(* IEC 61131-3 sources: test/Class/SdiasSDCIMaster (part 4) *)

          GetSdoReadData(pLength:=#TempDataLen, pData:=#TempData[0]);
          if TempDataLen = 9 then
            // check response data
            if (TempData[0] = (E_FNCID_CNTSTA)$USINT) then // check function ID
              // reset response state machine
              sSdoData.eResponseState := t_ReponseState::_PrepareSendData;

              // if the operating flags are cleared we can continue
              for i:= 0 to SIOL_MAX_PORTS_SUPPORTED-1 do
                TempStateFlags := TempData[1 + i*sizeof(t_StatusFlags)]$t_StatusFlags;

                // if any operating bit of the SDCI ports is still set and we did not exceed the timeout => go to wait for disabled
                if (aPortInfo[i].CfgPortMode = _SDCI) & (TempStateFlags.Operating = TRUE) &
                   ((ops.tAbsolute - Wait4DeviceDisableStartTime) < aPortInfo[sSdoData.ActPortSelection].udModeChangeTime) then

                  sSdoData.eInitSSW   := t_InitSSW::_Wait4DisableMode2;
                  return;
                end_if;
              end_for;

              // finished, continue with next step
              sSdoData.eInitSSW   := t_InitSSW::_Configure2StartUpMode;

            else
              // unexpected answer data
              LogError("@0525 (SdiasSDCIMaster::InitTheModule) Unexpected data in answer from µC: wrong function ID or port number (_SwitchToDisableMode2)");
              sSdoData.eInitSSW := _Error;
              return;
            end_if;
          else
            // invalid length of answer data
            LogError("@0526 (SdiasSDCIMaster::InitTheModule) Invalid data length in answer from µC (_SwitchToDisableMode2)");
            sSdoData.eInitSSW := _Error;
            return;
          end_if;

      //***************************************************************************************************
      end_case;

//**********************************************************************************************************************************************************
  	t_InitSSW::_Configure2StartUpMode:
      // if it's an SDCI port and physically available, we must wait the time (according to the specification), because some sensors might need it
      if (aPortInfo[sSdoData.ActPortSelection].CfgPortMode = _SDCI) &
          aPortInfo[sSdoData.ActPortSelection].PhysicallyAvailable  &
         ((ops.tAbsolute - Wait4DeviceDisableStartTime) < aPortInfo[sSdoData.ActPortSelection].udModeChangeTime) then
        return;
      end_if;

      case sSdoData.eResponseState of
      //***************************************************************************************************
        t_ReponseState::_PrepareSendData: // start the sending action

          // only if the port is of type SDCI and the device is physically available
          if (aPortInfo[sSdoData.ActPortSelection].CfgPortMode = _SDCI) & aPortInfo[sSdoData.ActPortSelection].PhysicallyAvailable &
             (aPortInfo[sSdoData.ActPortSelection].StartUpMode <> _Inactive) then

            // prepare the sdo buffer
            TempData[0]       := E_FNCID_SETPORTCNFPAR; // function ID
            TempData[1]       := sSdoData.ActPortSelection; // port number

            case aPortInfo[sSdoData.ActPortSelection].StartUpMode of
            //***************************************************************************************************
              _DigitalInput:
                TempData[2]       := t_OpModeStates::E_OPMODE_DI; // operating mode

            //***************************************************************************************************
              _DigitalOutput:
                TempData[2]       := t_OpModeStates::E_OPMODE_DO; // operating mode

            //***************************************************************************************************
              _SDCI:
                TempData[2]       := t_OpModeStates::E_OPMODE_FIXEDMODE; // operating mode

            //***************************************************************************************************
            end_case;

            TempData[3]       := t_PortCycle::E_PORTCYCLE_FIXVAL; // port cycle

            // check if a user override is active
            if aPortInfo[sSdoData.ActPortSelection].OverrideMinCycleTime_us then
              // recalculate cycle time from [µs] to [100µs]
              TempCycleTime     := to_uint(aPortInfo[sSdoData.ActPortSelection].OverrideMinCycleTime_us / 100);
            else
              // recalculate cycle time from [µs] to [100µs]
              TempCycleTime     := to_uint(aPortInfo[sSdoData.ActPortSelection].MinCycleTime_us / 100);
            end_if;

            // make endian swap
            TempCycleTime     := ((TempCycleTime SHR 8) AND 16#FF) OR ((TempCycleTime SHL 8) AND 16#FF00);

            TempData[4]$UINT  := TempCycleTime; // cycle time
            TempData[6]       :=  aPortInfo[sSdoData.ActPortSelection].PdoMapping.ReadDataLength$USINT; // PDConfig LenIn
            TempData[7]       := (aPortInfo[sSdoData.ActPortSelection].PdoMapping.ReadDataStartAddress - SIOL_OFFSET_RT_READ_DATA)$USINT; // PdConfig PosIn
            TempData[8]       := 0; // PdConfig SrcOffsetIn
            TempData[9]       :=  aPortInfo[sSdoData.ActPortSelection].PdoMapping.WriteDataLength$USINT; // PDConfig LenOut
            TempData[10]      := (aPortInfo[sSdoData.ActPortSelection].PdoMapping.WriteDataStartAddress - SIOL_OFFSET_RT_WRITE_DATA)$USINT; // PdConfig PosOut
            TempData[11]      := 0; // PdConfig SrcOffsetOut
            TempData[12]      := (aPortInfo[sSdoData.ActPortSelection].VendorID SHR 8)$USINT; // VendorID
            TempData[13]      :=  aPortInfo[sSdoData.ActPortSelection].VendorID$USINT; // VendorID
            TempData[14]      := (aPortInfo[sSdoData.ActPortSelection].DeviceID SHR 24)$USINT; // DeviceID
            TempData[15]      := (aPortInfo[sSdoData.ActPortSelection].DeviceID SHR 16)$USINT; // DeviceID
            TempData[16]      := (aPortInfo[sSdoData.ActPortSelection].DeviceID SHR  8)$USINT; // DeviceID
            TempData[17]      := (aPortInfo[sSdoData.ActPortSelection].DeviceID       )$USINT; // DeviceID
  //          _strcpy(dest:=#TempData[18], src:="0000000000000000"); // serial number as string
            _memset(dest:=#TempData[18], usByte:=0, cntr:=16); // serial number as string
            TempData[34]      := 1; // Inspection level (1 = device and vendor id have to match)
            TempData[35]      := 0; // DS activation state
            TempData[36]      := 0; // DS download enable
            TempData[37]      := 0; // DS upload enable
            TempData[38]      := aPortInfo[sSdoData.ActPortSelection].RevisionID; // revision ID

            TempDataLen := 39;

            InitializeSdoWriteData(Usage:=_SendFunctionCode, ParaIndex:=0, ParaSubIndex:=0, PortSelection:=SIOL_MASTER_PORT_NO, LengthOfData:=TempDataLen, pData:=#TempData[0]);

            sSdoData.eResponseState := t_ReponseState::_SendData;
          else
            if (aPortInfo[sSdoData.ActPortSelection].CfgPortMode = _SDCI) & (aPortInfo[sSdoData.ActPortSelection].StartUpMode = _Inactive) &
                aPortInfo[sSdoData.ActPortSelection].PhysicallyAvailable then
              // the current mode is now the startupmode
              aPortInfo[sSdoData.ActPortSelection].ActPortMode := aPortInfo[sSdoData.ActPortSelection].StartUpMode;

              // it's always ok here
              MyPara.aPara[0] := _ClassOk$DINT;

              // vendor ID
              MyPara.aPara[1] := aPortInfo[sSdoData.ActPortSelection].VendorID;

              // device ID
              MyPara.aPara[2] := aPortInfo[sSdoData.ActPortSelection].DeviceID$DINT;

              // minimum cycle time
              // check if a user override is active
              if aPortInfo[sSdoData.ActPortSelection].OverrideMinCycleTime_us then
                MyPara.aPara[3] := aPortInfo[sSdoData.ActPortSelection].OverrideMinCycleTime_us$DINT;
              else
                MyPara.aPara[3] := aPortInfo[sSdoData.ActPortSelection].MinCycleTime_us$DINT;
              end_if;

              // actual port mode is already valid here (no further changes on the setting of this port)
              MyPara.aPara[4] := aPortInfo[sSdoData.ActPortSelection].ActPortMode$DINT;

              aPortInfo[sSdoData.ActPortSelection].pThis^.NewInst(#MyPara, #MyResult);
            end_if;

            // already the last port?
            if sSdoData.ActPortSelection = (SIOL_MAX_PORTS_SUPPORTED-1) then
              // finished, continue with next step
              sSdoData.ActPortSelection := 0;
              DelayedEnablePorts        := 0;
              DigStartUpAvailable       := FALSE;

              for i:= 0 to SIOL_MAX_PORTS_SUPPORTED-1 do
                if (aPortInfo[i].CfgPortMode = _SDCI) & aPortInfo[i].PhysicallyAvailable then
                  if (aPortInfo[i].StartUpMode = _SDCI) then
                    DelayedEnablePorts := DelayedEnablePorts OR (1 SHL i$USINT);
                  elsif (aPortInfo[i].StartUpMode = _DigitalInput) | (aPortInfo[i].StartUpMode = _DigitalOutput) then
                    DigStartUpAvailable := TRUE;
                  end_if;
                end_if;
              end_for;

              if DelayedEnablePorts then
                // block the asynchron communication channel already
                sSdoData.AsyState             := t_SDCIRetCode::SDCI_Busy;
                sSdoData.TargetMode           := _SDCI;
                sSdoData.AsyCmdType           := t_AsyCmdType::DelayedEnable;
                sSdoData.eAsySSW              := t_AsySSW::_StartDelayedEnable;
                DelayedEnablePorts.FirstTime  := TRUE; // this is set to reset the port number on the first entrace in cyclic
              end_if;

              if DigStartUpAvailable then
                sSdoData.eInitSSW   := t_InitSSW::_EnableDigIOStartUpModes;
              else
                sSdoData.eInitSSW   := t_InitSSW::_SetCycleTimes;
              end_if;
            else
              // repeat the steps with the next port
              sSdoData.ActPortSelection += 1;
            end_if;
          end_if;

      //***************************************************************************************************
        t_ReponseState::_SendData,
        t_ReponseState::_Wait4SendResponse,
        t_ReponseState::_GotSendResponse,
        t_ReponseState::_ReadData,
        t_ReponseState::_Wait4ReceiveData,
        t_ReponseState::_GotReceiveData:
          if HandleSdoDataTransfer() = ERROR then
            sSdoData.eInitSSW := _Error;
            return;
          end_if;

      //***************************************************************************************************
        t_ReponseState::_GotAllReceiveData:// we enter this step, when we received the answer with the data

          GetSdoReadData(pLength:=#TempDataLen, pData:=#TempData[0]);
          if TempDataLen = 3 then
            // check response data
            if (TempData[0] = (E_FNCID_SETPORTCNFPAR)$USINT) & // check function ID
               (TempData[1] = sSdoData.ActPortSelection)              // check port number
               then

              if (TempData[2] = 0) then // check status code seperately
                // reset response state machine
                sSdoData.eResponseState := t_ReponseState::_PrepareSendData;

                // already the last port?
                if sSdoData.ActPortSelection = (SIOL_MAX_PORTS_SUPPORTED-1) then
                  // finished, continue with next step
                  sSdoData.ActPortSelection := 0;
                  DelayedEnablePorts        := 0;
                  DigStartUpAvailable       := FALSE;

                  for i:= 0 to SIOL_MAX_PORTS_SUPPORTED-1 do
                    if (aPortInfo[i].StartUpMode = _SDCI) & aPortInfo[i].PhysicallyAvailable then
                      DelayedEnablePorts := DelayedEnablePorts OR (1 SHL i$USINT);
                    elsif (aPortInfo[i].CfgPortMode = _SDCI)         &  aPortInfo[i].PhysicallyAvailable &
                         ((aPortInfo[i].StartUpMode = _DigitalInput) | (aPortInfo[i].StartUpMode = _DigitalOutput)) then
                      DigStartUpAvailable := TRUE;
                    end_if;
                  end_for;

                  if DelayedEnablePorts then
                    // block the asynchron communication channel already
                    sSdoData.AsyState             := t_SDCIRetCode::SDCI_Busy;
                    sSdoData.TargetMode           := _SDCI;
                    sSdoData.AsyCmdType           := t_AsyCmdType::DelayedEnable;
                    sSdoData.eAsySSW              := t_AsySSW::_StartDelayedEnable;
                    DelayedEnablePorts.FirstTime  := TRUE; // this is set to reset the port number on the first entrace in cyclic
                  end_if;

                  if DigStartUpAvailable then
                    sSdoData.eInitSSW   := t_InitSSW::_EnableDigIOStartUpModes;
                  else
                    sSdoData.eInitSSW   := t_InitSSW::_SetCycleTimes;
                  end_if;
                else
                  // repeat the steps with the next port
                  sSdoData.ActPortSelection += 1;
                end_if;
              else
                // error at return code
                LogError("@0527 (SdiasSDCIMaster::InitTheModule) Error at status code in answer from µC (_Configure2StartUpMode)");
                sSdoData.eInitSSW := _Error;
                return;
              end_if;
            else
              // unexpected answer data
              LogError("@0529 (SdiasSDCIMaster::InitTheModule) Unexpected data in answer from µC: wrong function ID or port number (_ReEnableWithFixedMode)");
              sSdoData.eInitSSW := _Error;
              return;
            end_if;
          else
            // invalid length of answer data
            LogError("@052A (SdiasSDCIMaster::InitTheModule) Invalid data length in answer from µC (_Configure2StartUpMode)");
            sSdoData.eInitSSW := _Error;
            return;
          end_if;

      //***************************************************************************************************
      end_case;

//**********************************************************************************************************************************************************
  	t_InitSSW::_EnableDigIOStartUpModes:
      case sSdoData.eResponseState of
      //***************************************************************************************************
        t_ReponseState::_PrepareSendData: // start the sending action
          TempFlags := 0;
          TempFlags.Start2Operate := TRUE;
          TempFlags.OperatingMode := TRUE;

          // prepare the sdo buffer
          TempData[0]       := E_FNCID_CNTSTA; // function ID
          for i:= 0 to SIOL_MAX_PORTS_SUPPORTED-1 do

            // if the startup mode is digin or digout => enable this mode now
            if (aPortInfo[i].CfgPortMode = _SDCI)         &  aPortInfo[i].PhysicallyAvailable &
              ((aPortInfo[i].StartUpMode = _DigitalInput) | (aPortInfo[i].StartUpMode = _DigitalOutput)) then
              TempData[1 + i*sizeof(UINT)]$UINT := TempFlags;
            else
              // otherwise don't do anything at this port
              TempData[1 + i*sizeof(UINT)]$UINT := 0;
            end_if;
          end_for;

          if TotalMappingWriteSize then
            _memset(dest:=#TempData[9], usByte:=0, cntr:=TotalMappingWriteSize);
          end_if;

          TempDataLen := 9 + TotalMappingWriteSize;

          InitializeSdoWriteData(Usage:=_SendFunctionCode, ParaIndex:=0, ParaSubIndex:=0, PortSelection:=SIOL_MASTER_PORT_NO, LengthOfData:=TempDataLen, pData:=#TempData[0]);

          sSdoData.eResponseState := t_ReponseState::_SendData;

      //***************************************************************************************************
        t_ReponseState::_SendData,
        t_ReponseState::_Wait4SendResponse,
        t_ReponseState::_GotSendResponse,
        t_ReponseState::_ReadData,
        t_ReponseState::_Wait4ReceiveData,
        t_ReponseState::_GotReceiveData:
          if HandleSdoDataTransfer() = ERROR then
            sSdoData.eInitSSW := _Error;
            return;
          end_if;

      //***************************************************************************************************
        t_ReponseState::_GotAllReceiveData:// we enter this step, when we received the answer with the data

          GetSdoReadData(pLength:=#TempDataLen, pData:=#TempData[0]);
          if TempDataLen = 9 then

            // reset response state machine
            sSdoData.eResponseState := t_ReponseState::_PrepareSendData;

            // check response data
            if (TempData[0] = (E_FNCID_CNTSTA)$USINT) then // check function ID

              // update the state of the object
              for i:= 0 to SIOL_MAX_PORTS_SUPPORTED-1 do

                // if the startup mode is digin or digout => show classok and current mode
                if (aPortInfo[i].CfgPortMode = _SDCI)         &  aPortInfo[i].PhysicallyAvailable
                & ((aPortInfo[i].StartUpMode = _DigitalInput) | (aPortInfo[i].StartUpMode = _DigitalOutput))
                  then
                  // the current mode is now the startupmode
                  aPortInfo[i].ActPortMode := aPortInfo[i].StartUpMode;

                  // it's always ok here
                  MyPara.aPara[0] := _ClassOk$DINT;

                  // vendor ID
                  MyPara.aPara[1] := aPortInfo[i].VendorID;

                  // device ID
                  MyPara.aPara[2] := aPortInfo[i].DeviceID$DINT;

                  // minimum cycle time
                  // check if a user override is active
                  if aPortInfo[i].OverrideMinCycleTime_us then
                    MyPara.aPara[3] := aPortInfo[i].OverrideMinCycleTime_us$DINT;
                  else
                    MyPara.aPara[3] := aPortInfo[i].MinCycleTime_us$DINT;
                  end_if;

                  // actual port mode is already valid here (no further changes on the setting of this port)
                  MyPara.aPara[4] := aPortInfo[i].ActPortMode$DINT;

                  aPortInfo[i].pThis^.NewInst(#MyPara, #MyResult);
                end_if;
              end_for;

              // finished, continue with next step
              sSdoData.eInitSSW   := t_InitSSW::_SetCycleTimes;

            else
              // unexpected answer data
              LogError("@050C (SdiasSDCIMaster::InitTheModule) Unexpected data in answer from µC: wrong function ID or port number (_SwitchToNewMode)");
              sSdoData.eInitSSW := _Error;
              return;
            end_if;
          else
            // invalid length of answer data
            LogError("@050D (SdiasSDCIMaster::InitTheModule) Invalid data length in answer from µC (_SwitchToNewMode)");
            sSdoData.eInitSSW := _Error;
            return;
          end_if;

      //***************************************************************************************************
      end_case;

//**********************************************************************************************************************************************************
  	t_InitSSW::_SetCycleTimes:

      case sSdoData.eResponseState of
      //***************************************************************************************************
        t_ReponseState::_PrepareSendData: // start the sending action

          // take the time from the parameter download process
          ParaDownloadTime := ops.tAbsolute - DownloadTimeStart;

          TempData[0]$UINT  := (udBusTime / 1000)$UINT; // SDIAS Bus cycle time
          TempData[2]$UINT  := CycleTime$UINT;

          TempDataLen    := 2 * sizeof(UINT);

          InitializeSdoWriteData(Usage:=_SendCycleTimeInfo, ParaIndex:=0, ParaSubIndex:=0, PortSelection:=SIOL_MASTER_PORT_NO, LengthOfData:=TempDataLen, pData:=#TempData[0]);

          sSdoData.eResponseState := t_ReponseState::_SendData;

      //***************************************************************************************************
        t_ReponseState::_SendData,
        t_ReponseState::_Wait4SendResponse,
        t_ReponseState::_GotSendResponse,
        t_ReponseState::_ReadData,
        t_ReponseState::_Wait4ReceiveData,
        t_ReponseState::_GotReceiveData:
          if HandleSdoDataTransfer() = ERROR then
            sSdoData.eInitSSW := _Error;
            return;
          end_if;

      //***************************************************************************************************
        t_ReponseState::_GotAllReceiveData:// we enter this step, when we received the answer with the data

          GetSdoReadData(pLength:=#TempDataLen, pData:=#TempData[0]);
          if TempDataLen = 0 then
            // check response data
            if (sSdoData.SdoReadData.ro_RetCode = _FwOk) then // check returncode
              // reset response state machine
              sSdoData.eResponseState := t_ReponseState::_SendData;

              sSdoData.RemainingDataSize := SIOL_MAX_PORTS_SUPPORTED * SIOL_MAX_PDO_SIZE;
              sSdoData.ActDataSize       := SDIAS_MAX_SDO_WRITE_LENGTH;
              sSdoData.pActData          := #LocalWritePDOBuf;

              // finished, continue with next step
              sSdoData.eInitSSW   := t_InitSSW::_ResetOutputImage;
            else
              // error
              LogError("@052A (SdiasSDCIMaster::InitTheModule) Error reported by µC (_SetCycleTimes)");
              sSdoData.eInitSSW := _Error;
              return;
            end_if;
          else
            // invalid length of answer data
            LogError("@052B (SdiasSDCIMaster::InitTheModule) Invalid data length in answer from µC (_SetCycleTimes)");
            sSdoData.eInitSSW := _Error;
            return;
          end_if;

      //***************************************************************************************************
      end_case;

//**********************************************************************************************************************************************************
  	t_InitSSW::_ResetOutputImage:
      case sSdoData.eResponseState of
        //***************************************************************************************************
          t_ReponseState::_SendData:// we enter this step to start the read access

            StartWriteSDO(hOffset:=SIOL_OFFSET_RT_WRITE_DATA, usLength:=sSdoData.ActDataSize, pWriteBuffer:=sSdoData.pActData$^USINT, eCommand:=SDIAS_SDO_CMD_MEM_WRITE);

            sSdoData.TimeoutStart   := ops.tAbsolute;
            sSdoData.eResponseState := t_ReponseState::_Wait4SendResponse;

        //***************************************************************************************************
          t_ReponseState::_Wait4SendResponse:// we wait for the read data
            if (ops.tAbsolute - sSdoData.TimeoutStart) > SIOL_SDO_TIMEOUT then
              LogError("@052C (SdiasSDCIMaster::InitTheModule) Timeout at resetting output image at module");
              sSdoData.eInitSSW := _Error;
              return;
            end_if;

        //***************************************************************************************************
          t_ReponseState::_GotSendResponse:// we enter this step, when we received the answer with the data

            // here we decide if more packages need to be sent
            sSdoData.RemainingDataSize -= sSdoData.ActDataSize;
            sSdoData.pActData          += sSdoData.ActDataSize;

            if sSdoData.RemainingDataSize then
              // another write access is necessary, prepare the variables
              if sSdoData.RemainingDataSize > SDIAS_MAX_SDO_WRITE_LENGTH then
                // limit the act size to it's maximum
                sSdoData.ActDataSize := SDIAS_MAX_SDO_WRITE_LENGTH;
              else
                // last package
                sSdoData.ActDataSize := sSdoData.RemainingDataSize;
              end_if;

              // send the next package
              sSdoData.eResponseState := t_ReponseState::_SendData;
            else
              // finished with writing => go to reading the answer
              sSdoData.eResponseState   := t_ReponseState::_PrepareSendData;
              sSdoData.eInitSSW   := t_InitSSW::_Finished;
            end_if;

        //***************************************************************************************************
      end_case;

//**********************************************************************************************************************************************************
  	t_InitSSW::_Finished:

      // Enable Buffer
      HWKVarSizeFIFO1.Enable();

      // Unlock SDO Channel
      sigclib_atomic_setU32(pValue:=#sSdoData.DataLock, value:= SSDCIM_SDO_UNLOCK);

      eModuleInitState := READY;
      eInitState       := _ClassOk;

//**********************************************************************************************************************************************************
  	t_InitSSW::_Error:

      // Do not unlock SDO Channel module is not working!
      eModuleInitState := ERROR;
      if eInitState = _NotInitialized then
        eInitState    := _InvalidConfguration;
      end_if;

//**********************************************************************************************************************************************************
  end_case;

#ifdef SIOL_ENABLE_DEBUG_LOGGING
  if sSdoData.eInitSSW <> OldStep then
    StepTimes[OldStep$DINT] := ops.tAbsolute;
    OldStep := sSdoData.eInitSSW;
  end_if;
#pragma message("RamAnd 31.01.2017 10:41 \ testweise die Zeit der einzelnen Steps messen")
#endif

END_FUNCTION

FUNCTION VIRTUAL SdiasSDCIMaster::HandleSDOFifo
  VAR
  	localSDOLock : UDINT;
    datasize : DINT;
    sSDOFIFOHeader : t_SDOFIFOHeader;
    aDatatmp    : array [0..SIOL_MAX_SDO_DATA_SIZE - 1] of USINT;
    bEndianSwapNeeded : BOOL;
    pParaInfo   : ^t_ConfigTablePara;
  END_VAR

  localSDOLock := sigclib_atomic_cmpxchgU32(pValue:=#sSdoData.DataLock, cmpVal := SSDCIM_SDO_UNLOCK, newVal := SSDCIM_SDO_LOCK);

  // Get Lock on SDO Channel
  if localSDOLock = SSDCIM_SDO_UNLOCK then

    // Get next sSDOFIFOHeader from buffer
    datasize := HWKVarSizeFIFO1.ReadData(pData := (#sSDOFIFOHeader)$^HSINT, size := sizeof(sSDOFIFOHeader));

    // Check if header is valid
    if datasize = sizeof(sSDOFIFOHeader) then

      // Always safe callback pointers
      sSdoData.pCallBackThis  := sSDOFIFOHeader.pThis;
      sSdoData.pCallBackFun   := sSDOFIFOHeader.pCallBackFunction;

      case sSDOFIFOHeader.NewInstCmd of

//**********************************************************************************************************************************************************
        CMD_SIOL_DEVICE_SET_PORT_MODE_BUFFERED:

          sSdoData.ActPortSelection := sSDOFIFOHeader.PortSelection;

          datasize := HWKVarSizeFIFO1.GetData(pData   := (#sSdoData.TargetMode)$^HSINT
                                            , size    := sizeof(t_SDCIPortMode)
                                            , offset  := sizeof(sSDOFIFOHeader));

          if (datasize <> sizeof(t_SDCIPortMode) ) then

            LogValue(pString := "@052D (SdiasSDCIMaster::HandleSDOFifo) Invalid LengthOfData 0x{0} in Fifo, Command = 0x{1}", udValue:=datasize$UDINT, udValue2:= sSDOFIFOHeader.NewInstCmd);
            // Unlock SDO Channel
            sigclib_atomic_setU32(pValue:=#sSdoData.DataLock, value:= SSDCIM_SDO_UNLOCK);
            return;

//          else
//            // Data Ok
          end_if;

          // we're busy now
          sSdoData.AsyState         := t_SDCIRetCode::SDCI_Busy;

          sSdoData.AsyCmdType       := t_AsyCmdType::ModeChange;
          sSdoData.eAsySSW          := t_AsySSW::_StartModeChange;
          sSdoData.eResponseState   := t_ReponseState::_SendData;
          sSdoData.AsyErrorCode     := t_SDCIRetCode::SDCI_UnspecifiedError;

//**********************************************************************************************************************************************************
        CMD_SIOL_DEVICE_RECONNECT_BUFFERED:

          // we're busy now
          sSdoData.AsyState         := t_SDCIRetCode::SDCI_Busy;

          sSdoData.ActPortSelection := sSDOFIFOHeader.PortSelection;

          sSdoData.AsyCmdType       := t_AsyCmdType::Reconnect;
          sSdoData.eAsySSW          := t_AsySSW::_StartReconnect;
          sSdoData.eResponseState   := t_ReponseState::_SendData;
          sSdoData.AsyErrorCode     := t_SDCIRetCode::SDCI_UnspecifiedError;

          HWKVarSizeFIFO1.RemoveData();

//**********************************************************************************************************************************************************
        CMD_SIOL_DEVICE_GET_ASY_PARA_BUFFERED,
        CMD_SIOL_DEVICE_SET_ASY_PARA_BUFFERED,
        CMD_SIOL_DEVICE_ASY_FUNCTION_ID_BUFFERED:

            // reset some parts of the readdata structure
            sSdoData.SdoReadData.ro_Checksum    := 0;

            // initialize variables for the cyclic state machine
            sSdoData.SdoWriteData.ParaIndex     := sSDOFIFOHeader.ParaIndex;
            sSdoData.SdoWriteData.ParaSubIndex  := sSDOFIFOHeader.ParaSubIndex;
            sSdoData.SdoWriteData.PortSelection := sSDOFIFOHeader.PortSelection;
            sSdoData.SdoWriteData.LengthOfData  := sSDOFIFOHeader.LengthOfData;

            if sSdoData.SdoWriteData.LengthOfData then

              if sSdoData.SdoWriteData.LengthOfData <= SIOL_MAX_SDO_DATA_SIZE then

                // Get the infomation bEndianSwapNeeded
                bEndianSwapNeeded := FALSE;
                if ( sSdoData.SdoWriteData.PortSelection < SIOL_MAX_PORTS_SUPPORTED) then

                  // Get parameter information
                  pParaInfo := FindParaInTable( pActPortInfo := #aPortInfo[sSdoData.SdoWriteData.PortSelection]
                                              , ParaID       := sSdoData.SdoWriteData.ParaIndex
                                              , ParaSubID    := sSdoData.SdoWriteData.ParaSubIndex);

                  // Check if parameter needes endianswap
                  bEndianSwapNeeded := CheckEndianSwapNeeded( pParaInfo     := pParaInfo
                                                            , PortSelection := sSdoData.SdoWriteData.PortSelection);
                end_if;

                if ( bEndianSwapNeeded = TRUE) then

                  // Get temp write data directly from buffer
                  datasize := HWKVarSizeFIFO1.GetData(  pData   := #aDatatmp[0]
                                                      , size    := sSdoData.SdoWriteData.LengthOfData
                                                      , offset  := sizeof(sSDOFIFOHeader));

                  if (datasize = sSdoData.SdoWriteData.LengthOfData) then
                    // Endianswap write data
                    EndianSwap( pDst          := #sSdoData.SdoWriteData.aData[SIOL_MAX_SDO_DATA_SIZE-sSdoData.SdoWriteData.LengthOfData]
                              , pSrc          := #aDatatmp[0]
                              , LengthOfData  := sSdoData.SdoWriteData.LengthOfData);
                  // else
                  //   LogValue(pString := "@052D (SdiasSDCIMaster::HandleSDOFifo) Invalid LengthOfData 0x{0} in Fifo, Command = 0x{1}", udValue:=datasize$UDINT, udValue2:= sSDOFIFOHeader.NewInstCmd);
                  end_if;

                else
                  // Get write data directly from buffer
                  datasize := HWKVarSizeFIFO1.GetData(  pData   := #sSdoData.SdoWriteData.aData[SIOL_MAX_SDO_DATA_SIZE-sSdoData.SdoWriteData.LengthOfData]
                                                      , size    := sSdoData.SdoWriteData.LengthOfData
                                                      , offset  := sizeof(sSDOFIFOHeader));
                end_if;

                if (datasize <> sSdoData.SdoWriteData.LengthOfData) then

                  LogValue(pString := "@052D (SdiasSDCIMaster::HandleSDOFifo) Invalid LengthOfData 0x{0} in Fifo, Command = 0x{1}", udValue:=datasize$UDINT, udValue2:= sSDOFIFOHeader.NewInstCmd);
                  // Unlock SDO Channel
                  sigclib_atomic_setU32(pValue:=#sSdoData.DataLock, value:= SSDCIM_SDO_UNLOCK);
                  return;

      //          else
      //            // Data Ok
                end_if;

              else
                LogValue(pString := "@052D (SdiasSDCIMaster::HandleSDOFifo) Invalid LengthOfData 0x{0} in Fifo, Command = 0x{1}", udValue:=datasize$UDINT, udValue2:= sSDOFIFOHeader.NewInstCmd);

                // Remove Invalid Data from Fifo
                HWKVarSizeFIFO1.RemoveData();
                // Unlock SDO Channel
                sigclib_atomic_setU32(pValue:=#sSdoData.DataLock, value:= SSDCIM_SDO_UNLOCK);
                return;
              end_if;
            else
              HWKVarSizeFIFO1.RemoveData();
            end_if;

            case sSDOFIFOHeader.NewInstCmd of

              CMD_SIOL_DEVICE_GET_ASY_PARA_BUFFERED:

                sSdoData.SdoWriteData.wo_ActUsage   := _ReadParaData;

              CMD_SIOL_DEVICE_SET_ASY_PARA_BUFFERED:

                sSdoData.SdoWriteData.wo_ActUsage   := _WriteParaData;

              CMD_SIOL_DEVICE_ASY_FUNCTION_ID_BUFFERED:

                sSdoData.SdoWriteData.wo_ActUsage   := _SendFunctionCode;

            end_case;

            sSdoData.SdoWriteData.wo_MessageCnt += 1;
            sSdoData.SdoWriteData.wo_Checksum   := CalcChecksum(Mode:=1);

            // set RemainingDataSize, pActData and ActDataSize correctly for the first send package

            // at the initialisation we set the remaining size to the complete package that needs to be transferred
            sSdoData.RemainingDataSize  := sSdoData.SdoWriteData.LengthOfData + sizeof(t_ServiceDataArea) - sizeof(t_ServiceDataArea.aData) - sizeof(t_ServiceDataArea.ro_MessageCnt) - sizeof(t_ServiceDataArea.ro_RetCode) - sizeof(t_ServiceDataArea.ro_Checksum);
            sSdoData.pActData           := #sSdoData.SdoWriteData + SIOL_MAX_SDO_DATA_SIZE - sSdoData.SdoWriteData.LengthOfData;
            if sSdoData.RemainingDataSize > SDIAS_MAX_SDO_WRITE_LENGTH then
              // limit the act size to it's maximum
              sSdoData.ActDataSize := SDIAS_MAX_SDO_WRITE_LENGTH;
            else
              // we only need one package
              sSdoData.ActDataSize := sSdoData.RemainingDataSize;
            end_if;

            sSdoData.AsyState       := t_SDCIRetCode::SDCI_Busy;
            sSdoData.AsyCmdType     := t_AsyCmdType::SingleAsyTransfer;
            sSdoData.eResponseState := t_ReponseState::_SendData;

//**********************************************************************************************************************************************************
      else
        LogValue("@04FB (SdiasSDCIMaster::HandleSDOFifo) Invalid command: 0x{0}" , udValue:= sSDOFIFOHeader.NewInstCmd);

        // Remove Invalid Data from Fifo
        HWKVarSizeFIFO1.RemoveData();
        // Unlock SDO Channel
        sigclib_atomic_setU32(pValue:=#sSdoData.DataLock, value:= SSDCIM_SDO_UNLOCK);
        return;
      end_case;

    else
      // No data in FIFO
      // Unlock SDO Channel
      sigclib_atomic_setU32(pValue:=#sSdoData.DataLock, value:= SSDCIM_SDO_UNLOCK);
    end_if;

//  else
//    // SDO Channel busy, do nothing
  end_if;

END_FUNCTION

FUNCTION VIRTUAL SdiasSDCIMaster::HandleSDOCallback
  VAR
  	AsyStatetmp : t_SDCIRetCode;
    pDatatmp    : ^USINT;
    bEndianSwapNeeded : BOOL;
    pParaInfo   : ^t_ConfigTablePara;
  END_VAR

  AsyStatetmp := sSdoData.AsyState;
  pDatatmp    := NIL;

  if (sSdoData.SdoReadData.LengthOfData) then

    if (sSdoData.SdoReadData.LengthOfData <= SIOL_MAX_SDO_DATA_SIZE) then

      // Get the infomation bEndianSwapNeeded
      bEndianSwapNeeded := FALSE;
      if ( sSdoData.SdoReadData.PortSelection < SIOL_MAX_PORTS_SUPPORTED) then

        // Get parameter information
        pParaInfo := FindParaInTable( pActPortInfo := #aPortInfo[sSdoData.SdoReadData.PortSelection]
                                    , ParaID       := sSdoData.SdoReadData.ParaIndex
                                    , ParaSubID    := sSdoData.SdoReadData.ParaSubIndex);

        // Check if parameter needes endianswap
        bEndianSwapNeeded := CheckEndianSwapNeeded( pParaInfo     := pParaInfo
                                                  , PortSelection := sSdoData.SdoReadData.PortSelection);
      end_if;

      if bEndianSwapNeeded = TRUE then
        EndianSwap( pDst          := #sSdoData.SdoReadDataSwapped[SIOL_MAX_SDO_DATA_SIZE-sSdoData.SdoReadData.LengthOfData]
                  , pSrc          := #sSdoData.SdoReadData.aData[SIOL_MAX_SDO_DATA_SIZE-sSdoData.SdoReadData.LengthOfData]
                  , LengthOfData  := sSdoData.SdoReadData.LengthOfData);

        // Pass pointer to swapped data
        pDatatmp := #sSdoData.SdoReadDataSwapped[SIOL_MAX_SDO_DATA_SIZE-sSdoData.SdoReadData.LengthOfData];

      else

        // Pass pointer to data
        pDatatmp := #sSdoData.SdoReadData.aData[SIOL_MAX_SDO_DATA_SIZE-sSdoData.SdoReadData.LengthOfData];
      end_if;

    else
      AsyStatetmp := t_SDCIRetCode::SDCI_MicroCtrl_RspLengthTooBig;
    end_if;

  end_if;

  sSdoData.pCallBackFun$AsyCallBackSdiasSDCIMaster( pThis         := sSdoData.pCallBackThis
                                                  , AsyState      := AsyStatetmp
                                                  , LengthOfData  := sSdoData.SdoReadData.LengthOfData
                                                  , pData         := pDatatmp);

  // Don't care about return code. If reciever can't handle callback that's his problem.

END_FUNCTION

FUNCTION VIRTUAL SdiasSDCIMaster::CheckEndianSwapNeeded
	VAR_INPUT
		pParaInfo 	  : ^t_ConfigTablePara;
    PortSelection : USINT;
	END_VAR
	VAR_OUTPUT
		bCheckEndianSwapNeeded 	: BOOL;
	END_VAR

  bCheckEndianSwapNeeded := FALSE;

  if ( (PortSelection < SIOL_MAX_PORTS_SUPPORTED) &
       (aPortInfo[PortSelection].SkipEndianSwapAsy = FALSE) ) then

    if pParaInfo then

      // Swap is only needed for _Float32, _Int16, _Int32, _Int64, _Uint16, _Uint32, _Uint64
      // Not needed for _Text and 1 Byte Parameters
      case pParaInfo^.DataType of

        _Float32,
        _Int16,
        _Int32,
        _Int64,
        _Uint16,
        _Uint32,
        _Uint64:
          bCheckEndianSwapNeeded := TRUE;

      end_case;

    end_if;
  end_if;

END_FUNCTION

FUNCTION SdiasSDCIMaster::EndianSwap
	VAR_INPUT
		pDst 	: ^USINT;
		pSrc 	: ^USINT;
		LengthOfData 	: USINT;
	END_VAR
  VAR
  	pDataSrc : ^USINT;
    pDataDst : ^USINT;
    i : DINT;
  END_VAR

  // Method can't handle pDst = pSrc
  if pDst & pSrc & LengthOfData & pDst <> pSrc then

    pDataSrc := pSrc + LengthOfData - 1;
    pDataDst := pDst;

    for i := 1 to LengthOfData do

      pDataDst^ := pDataSrc^;

      pDataSrc -= 1;
      pDataDst += 1;

    end_for;

  end_if;

END_FUNCTION

FUNCTION SdiasSDCIMaster::HandleAutoConnect
	VAR_INPUT
		usPortNbr 	: USINT;
	END_VAR
	VAR_OUTPUT
		retcode 	: SdiasSDCIMaster::t_SDCIRetCode;
	END_VAR
  VAR
  	udTimeDiff    : UDINT;
  	MyPara        : CmdStruct;
    MyResult      : results;
  END_VAR

  //initialize return code
  retcode := SdiasSDCIMaster::t_SDCIRetCode::SDCI_Ready_Ok;

  //check for valid port numbers
  if usPortNbr >= SIOL_MAX_PORTS_SUPPORTED then
    return;
  end_if;

  //if port is not configured for SDCI Device dont start port scan
  if aPortInfo[usPortNbr].StartUpMode <> _SDCI & aPortInfo[usPortNbr].ActPortMode <> _SDCI then
    return;
  end_if;

  //check asy read timeout of other asy accesses
  if sSdoData.bSingleAsyTransferReady = TRUE & (ops.tAbsolute-sSdoData.udSingleAsyTransferReady >= SIOL_TIMEOUT_GETASYNCHRONOUS_DATA) then
    //reset flag
    sSdoData.bSingleAsyTransferReady := FALSE;
  end_if;

  //check last reconnect time to allow other asy communication (SDCIDevice_AsyncPara) and wait for other asy accesses to get their data
  if (ops.tAbsolute-sAutoConnectVars.udLastReconnectTry) < WaitTimeReconnect (*SIOL_MINIMUM_wAIT4RECONNECT_TIME*)
  | (sSdoData.bSingleAsyTransferReady = TRUE) then
    retcode := SdiasSDCIMaster::t_SDCIRetCode::SDCI_Busy;
    return;
  end_if;

  //get act port timediff as ms
  udTimeDiff := (ops.tAbsolute - aPortInfo[usPortNbr].udStartConnect);
  //check if auto connect is enabled and interval time is reached for this port
  if aPortInfo[usPortNbr].PhysicallyAvailable = FALSE
  & aPortInfo[usPortNbr].udAutoConnectTime
  & aPortInfo[usPortNbr].udAutoConnectTime <= udTimeDiff then
    // set reconnect for this port to check for connected devices
    MyPara.uiCmd   := CMD_SIOL_DEVICE_RECONNECT;
    // add the port in the last parameter
    MyPara.aPara[MAXCMDPARA-1] := usPortNbr;

    MyResult.uiLng := 0;

    ClassState.NewInst(#MyPara, #MyResult);

    if MyResult.uiLng >= sizeof(SdiasSDCIMaster::t_SDCIRetCode) then
      retcode := MyResult.aData$SdiasSDCIMaster::t_SDCIRetCode;
    else
      retcode := SdiasSDCIMaster::t_SDCIRetCode::SDCI_UnspecifiedError;
    end_if;

    //if ok then reconnect is started
    if retcode = SDCI_Ready_Ok then
      //save timediff of reconnecting
      aPortInfo[usPortNbr].udStartConnTimeDiff := ops.tAbsolute - aPortInfo[usPortNbr].udStartConnect;
      //set last reconnect time stamp for wait time
      aPortInfo[usPortNbr].udStartConnect := ops.tAbsolute;
      sAutoConnectVars.bReConnectStarted := TRUE;
    end_if;
  end_if;

END_FUNCTION

FUNCTION TAB SdiasSDCIMaster::BitMask

  0xFF$USINT, // special, all bits needed if rest of bits is 0
  0x01$USINT,
  0x03$USINT,
  0x07$USINT,
  0x0F$USINT,
  0x1F$USINT,
  0x3F$USINT,
  0x7F$USINT

END_FUNCTION
